PROGRAM MAIN
VAR
	Hoi : BOOL;
	Hallo : BOOL;
END_VAR

END_PROGRAM

(* stored: Version 1.1.0.1
   POU MAIN: Id {32777243-1886-4d57-92c0-558c01be997c}, SpecialFunc None *)
